// TIA Portal V21 export
// export: Created 2026-10-23T20:44:56.2213109Z, ExportSetting WithDefaults, DisplayName Totally Integrated Automation Portal, DisplayVersion V21 Update 1, DisplayName SINAMICS Startdrive Advanced, DisplayVersion V21 HF2, DisplayName SINAMICS Startdrive G110M, G120, G120C, G120D, G120P, G115D, DisplayVersion V21 HF2, DisplayName SINAMICS Startdrive G130, G150, S120, S150, G200, G220, S200, S210, S220, Innomotics MVD, DisplayVersion V21 HF2, DisplayName STEP 7 Professional, DisplayVersion V21 Update 1, DisplayName STEP 7 Safety, DisplayVersion V21, DisplayName Tech WebApplication, DisplayVersion V21, DisplayName WinCC Basic/Comfort/Advanced, DisplayVersion V21 Update 1, DisplayName WinCC Unified, DisplayVersion V21 Update 1
TYPE "UDT_Motor_B16"
TITLE = Motor data
// stored: IsFailsafeCompliant false
   STRUCT
      Enable : Bool;   // Release from the line control
      Running : Bool;   // Feedback: motor is running
      Fault : Bool;   // Motor protection tripped
      SpeedSetpoint : Real := 1450.0;   // Speed setpoint in rpm
      ActualSpeed : Real;   // Measured speed in rpm
      RunTime : Time := T#0MS;   // Accumulated run time
      StartCount : DInt := 0;   // Number of starts
      Enable_1 : Bool;   // Duplicate member name
   END_STRUCT;
END_TYPE
